TYPE ST_EL3356CoeWriteData :
STRUCT
	wIdx: WORD;
	bySubIdx: BYTE;
	bWriteOK: BOOL;
	dwData: DWORD;
	nSize: UDINT;
END_STRUCT
END_TYPE

(* stored: Version 1.1.0.1, ProductVersion 3.1.4024.15
   DUT ST_EL3356CoeWriteData: Id {c9bf4766-9b06-412d-90c4-cfad2fe19631} *)
